DATA_BLOCK "SealedA"
{ S7_Optimized_Access := 'TRUE' }
VERSION : 0.1
NON_RETAIN
"Sealed"

BEGIN

END_DATA_BLOCK
